Fanuc KAREL source: kb00109.KL

-- PROVISIONAL review KL for V770-1; original PC SHA256 3ca94f93b59b369ad08c36e67f5d504f89142bbb4734ea8c47027f7d5d8f3474
-- Incomplete behavior may be omitted. Consult companion uncertainty JSON. Do not deploy.
PROGRAM KB00109
%NOLOCKGROUP
-- UNRESOLVED_DECL P1 type=000101
-- UNRESOLVED_DECL RESULT type=000101
BEGIN
  -- UNRESOLVED_PC offsets 5-32; opcodes 27,22,1C,76,7E,4A
  -- UNRESOLVED_PC offsets 37-41; opcodes 7F
END KB00109
